(* PLC project Vn_shl, Beckhoff Automation GmbH TwinCAT PLC Control 3.5.13.21 *)
(* stored: creationDateTime 1970-01-01T00:00:00 *)

PROGRAM Vn_shl

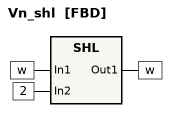
(* FBD diagram, written out as Structured Text *)
w := SHL(w, 2);
END_PROGRAM
